// TIA Portal project "Es02_Timer" (V18)

(* hardware
DEVICE "S71500/ET200MP station_1"  S7-1500 station
   slot 0: "Telaio di montaggio_0"  Rack  6ES7 590-1***0-0AA0
   slot 1: "PLC_1"  CPU 1516-3 PN/DP  6ES7 516-3AN01-0AB0  V2.5
      slot 3: "Display CPU_1"  6ES7591-1BA00-0AA0
   slot 2: "DI 32x24VDC HF_1"  DI 32x24VDC HF  6ES7 521-1BL00-0AB0  V2.1
   slot 3: "DQ 32x24VDC/0.5A HF_1"  DQ 32x24VDC/0.5A HF  6ES7 522-1BL01-0AB0  V1.0
   slot 4: "AI 8xU/I/RTD/TC ST_1"  AI 8xU/I/RTD/TC ST  6ES7 531-7KF00-0AB0  V2.1
   slot 5: "AQ 4xU/I ST_1"  AQ 4xU/I ST  6ES7 532-5HD00-0AB0  V2.1
*)

// ===== PLC "PLC_1"  CPU 1516-3 PN/DP =====

VAR_GLOBAL   // PLC tag table "Tabella delle variabili standard"
   "Led30" AT %Q3.0 : Bool;
   "Led31" AT %Q3.1 : Bool;
END_VAR

DATA_BLOCK "DB_Comandi"   // DB1
{ S7_Optimized_Access := 'TRUE' }
VERSION : 0.1
   VAR
      btnStart : Bool;
      btnStop : Bool;
   END_VAR
BEGIN
END_DATA_BLOCK

DATA_BLOCK "DB_Variabili"   // DB2
{ S7_Optimized_Access := 'TRUE' }
VERSION : 0.1
   VAR
      led30 : Bool;
      led31 : Bool;
      myTimerSTART : Bool;
      myTimerDONE : Bool;
      myTimerOUTPUT : Time;
      myTimerDURATA : Time;
      inEsecuzione : Bool;
   END_VAR
BEGIN
END_DATA_BLOCK

// folder: System blocks/Program resources

DATA_BLOCK "myTimer"   // DB3
{ S7_Optimized_Access := 'TRUE' }
AUTHOR : Simatic
FAMILY : IEC
NAME : IEC_TMR
VERSION : 1.0
// stored: InstanceOfName IEC_TIMER
"IEC_TIMER"
BEGIN
END_DATA_BLOCK

// folder: (top level)

FUNCTION "FC_Grafcet" : Void   // FC1, SCL
{ S7_Optimized_Access := 'TRUE' }
VERSION : 0.1
BEGIN
   // funzionamento: premendo btnStart il plc deve accendere i 2 led
   // dopo 5 secondi li deve spegnere
   // dopo altri 5 secondi riaccendere
   // fino a quando non premo btnStop
   // 
   // se premo btnStart avvio il timer
   IF "DB_Comandi".btnStart = TRUE THEN
       "DB_Variabili".inEsecuzione := TRUE;
       "DB_Variabili".myTimerSTART := TRUE;
       "DB_Comandi".btnStart := FALSE;
   END_IF;

   IF "DB_Comandi".btnStop = TRUE THEN
       "DB_Variabili".inEsecuzione := FALSE;
       "DB_Variabili".myTimerSTART := FALSE;
       "DB_Comandi".btnStop := FALSE;
   END_IF;
   // il funzionanmento ciclico del timer dipende dall variabile inEsecuzione
   IF "DB_Variabili".inEsecuzione = TRUE THEN
       "DB_Variabili".myTimerSTART := TRUE;
   ELSE
       "DB_Variabili".myTimerSTART := FALSE;
   END_IF;
   // gestisco il timer done (tick in c#)
   IF "DB_Variabili".inEsecuzione = TRUE AND "DB_Variabili".myTimerDONE = TRUE THEN
       // porto a FALSE, in modo tale che il timer possa ripartire
       // perchè altrimenti myTimerSTART già a TRUE e non viene sentita dal timer
       // idem il myTimerDONE sempre a TRUE non verrebbe gestito il DONE successivo
       "DB_Variabili".myTimerDONE := FALSE;
       "DB_Variabili".myTimerSTART := FALSE;
       //accendo/spengo i led
       "DB_Variabili".led30 := NOT "DB_Variabili".led30;
       "DB_Variabili".led31 := NOT "DB_Variabili".led31;
   END_IF;
END_FUNCTION

FUNCTION "FC_Timer" : Void   // FC2, SCL
{ S7_Optimized_Access := 'TRUE' }
VERSION : 0.1
BEGIN
   // imposto la durata del timer
   "DB_Variabili".myTimerDURATA := T#5s;
   // dichiaro (istanzio) il timer (trascino dalla schdea a destra temporizzatori)
   "myTimer".PT := "DB_Variabili".myTimerDURATA;
   "myTimer".TON(IN:="DB_Variabili".myTimerSTART,
                 PT:="DB_Variabili".myTimerDURATA,
                 Q=> "DB_Variabili".myTimerDONE,
                 ET=>"DB_Variabili".myTimerOUTPUT);
   // se non voglio passare i paramtrei nel costruttore, o dovessi variarli durante l'esecuzione posso
   // impostarli direttamente "myTimer".PT := "DB_Variabili".myTimerDURATA
END_FUNCTION

FUNCTION "FC_Uscite" : Void   // FC3, SCL
{ S7_Optimized_Access := 'TRUE' }
VERSION : 0.1
BEGIN
   // scrivo fisicamente le uscite
   // 
   // qui andranno inseriti gli eventuali controlli
   // di sicurezza (emergenza, protezioni, fotocellule)
   "Led30" := "DB_Variabili".led30;
   "Led31" := "DB_Variabili".led31;
END_FUNCTION

ORGANIZATION_BLOCK "Main"   // OB1, LAD, ProgramCycle
TITLE = "Main Program Sweep (Cycle)"
{ S7_Optimized_Access := 'TRUE' }
VERSION : 0.1
   VAR_INPUT
      Initial_Call : Bool;   // Initial call of this OB
      Remanence : Bool;   // =True, if remanent data are available
   END_VAR
   VAR_TEMP   // added for the SCL form of the ladder/FBD networks
      _w1 : Bool;
      _w2 : Bool;
   END_VAR
BEGIN

REGION Network 1
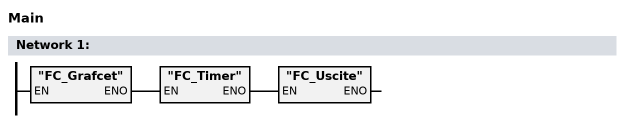
   RUNG wire#powerrail
      "FC_Grafcet"()
      "FC_Timer"()
      "FC_Uscite"()
   END_RUNG
   // the same network as SCL:
   "FC_Grafcet"(ENO => #_w1);
   "FC_Timer"(EN := #_w1, ENO => #_w2);
   IF #_w2 THEN "FC_Uscite"(); END_IF;
END_REGION
END_ORGANIZATION_BLOCK